Yaskawa INFORM job: LONGPRO5.JBI

/JOB
//NAME LONGPRO5
//POS
///NPOS 3,0,3,0,0,0
///TOOL 9
///POSTYPE PULSE
///PULSE
C00000=0,0,0
C00001=0,0,0
C00002=0,0,0
EC00000=0
EC00001=0
EC00002=0
//INST
<volatile>
///COMM Generated using RoboDK
///ATTR SC,RW
///GROUP1 RB1
NOP
MOVJ C00000 VJ=50.00  +MOVJ EC00000 VJ=100.00
MOVJ C00001 VJ=50.00  +MOVJ EC00001 VJ=100.00
MOVJ C00002 VJ=50.00  +MOVJ EC00002 VJ=100.00
END
